FUNCTION FC 1 : VOID
BEGIN
NETWORK
      A I 0.0
      XOR I 0.1
END_FUNCTION
